// TIA Portal V20 export
Screen "Pop-up_OPMode"  590x720
  ScreenItem "Rectangle TG1_14" at 21,669 size 548x40  Type=HmiRectangle
  ScreenItem "Rectangle TG1_13" at 21,628 size 548x40  Type=HmiRectangle
  ScreenItem "Rectangle TG1_12" at 21,588 size 548x40  Type=HmiRectangle
  ScreenItem "Rectangle TG1_11" at 21,548 size 548x40  Type=HmiRectangle
  ScreenItem "Rectangle TG1_10" at 21,508 size 548x40  Type=HmiRectangle
  ScreenItem "Rectangle TG1_9" at 21,467 size 548x40  Type=HmiRectangle
  ScreenItem "Background" at 21,65 size 548x32  Type=HmiRectangle
  ScreenItem "Rectangle TG1" at 21,101 size 548x40  Type=HmiRectangle
  ScreenItem "Text field TG1 Status" at 26,110 size 78x21  Type=HmiTextBox
  ScreenItem "Text field TG Status" at 1,0 size 589x47  Type=HmiTextBox
  ScreenItem "Rectangle TG1_1" at 21,141 size 548x40  Type=HmiRectangle
  ScreenItem "Text field TG1 Status_1" at 25,151 size 78x21  Type=HmiTextBox
  ScreenItem "Rectangle TG1_2" at 21,182 size 548x40  Type=HmiRectangle
  ScreenItem "Text field TG1 Status_2" at 25,187 size 78x21  Type=HmiTextBox
  ScreenItem "Rectangle TG1_3" at 21,222 size 548x40  Type=HmiRectangle
  ScreenItem "Text field TG1 Status_3" at 25,228 size 78x21  Type=HmiTextBox
  ScreenItem "Rectangle TG1_4" at 21,263 size 548x40  Type=HmiRectangle
  ScreenItem "Text field TG1 Status_4" at 25,271 size 78x21  Type=HmiTextBox
  ScreenItem "Rectangle TG1_5" at 21,304 size 548x40  Type=HmiRectangle
  ScreenItem "Text field TG1 Status_5" at 25,312 size 78x21  Type=HmiTextBox
  ScreenItem "Rectangle TG1_6" at 21,345 size 548x40  Type=HmiRectangle
  ScreenItem "Text field TG1 Status_6" at 26,352 size 78x21  Type=HmiTextBox
  ScreenItem "Rectangle TG1_7" at 21,385 size 548x40  Type=HmiRectangle
  ScreenItem "Text field TG1 Status_7" at 25,393 size 78x21  Type=HmiTextBox
  ScreenItem "Rectangle TG1_8" at 21,426 size 548x40  Type=HmiRectangle
  ScreenItem "Text field TG1 Status_8" at 25,435 size 78x21  Type=HmiTextBox
  ScreenItem "Text field TG1 Status_9" at 25,472 size 78x21  Type=HmiTextBox
  ScreenItem "Line_1" at 109,101 size 1x606  Type=HmiLine
  ScreenItem "Text field TG1 Status_10" at 115,111 size 440x21  Type=HmiTextBox
  ScreenItem "Text field TG1 Status_11" at 114,151 size 440x21  Type=HmiTextBox
  ScreenItem "Text field TG1 Status_12" at 114,189 size 440x21  Type=HmiTextBox
  ScreenItem "Text field TG1 Status_13" at 114,228 size 440x21  Type=HmiTextBox
  ScreenItem "Text field TG1 Status_14" at 114,270 size 440x21  Type=HmiTextBox
  ScreenItem "Text field TG1 Status_15" at 114,312 size 440x21  Type=HmiTextBox
  ScreenItem "Text field TG1 Status_16" at 115,351 size 440x21  Type=HmiTextBox
  ScreenItem "Text field TG1 Status_17" at 114,394 size 440x21  Type=HmiTextBox
  ScreenItem "Text field TG1 Status_18" at 114,436 size 440x21  Type=HmiTextBox
  ScreenItem "Text field TG1 Status_19" at 114,472 size 440x21  Type=HmiTextBox
  ScreenItem "Cancel Mode" at 505,3 size 82x42  Type=HmiButton
  ScreenItem "Text field TG1 Status_20" at 25,72 size 78x21  Type=HmiTextBox
  ScreenItem "Text field TG1 Status_21" at 218,72 size 260x21  Type=HmiTextBox
  ScreenItem "Text field TG1 Status_22" at 25,513 size 78x21  Type=HmiTextBox
  ScreenItem "Text field TG1 Status_23" at 114,513 size 440x21  Type=HmiTextBox
  ScreenItem "Text field TG1 Status_24" at 25,553 size 78x21  Type=HmiTextBox
  ScreenItem "Text field TG1 Status_25" at 114,553 size 440x21  Type=HmiTextBox
  ScreenItem "Text field TG1 Status_26" at 25,593 size 78x21  Type=HmiTextBox
  ScreenItem "Text field TG1 Status_27" at 114,593 size 440x21  Type=HmiTextBox
  ScreenItem "Text field TG1 Status_28" at 25,633 size 78x21  Type=HmiTextBox
  ScreenItem "Text field TG1 Status_29" at 114,633 size 440x21  Type=HmiTextBox
  ScreenItem "Text field TG1 Status_30" at 25,674 size 78x21  Type=HmiTextBox
  ScreenItem "Text field TG1 Status_31" at 114,674 size 440x21  Type=HmiTextBox
